// TIA Portal V20 export
TYPE "Stationsvariablen"
   STRUCT
      Anwahl_Tipp : Bool := FALSE;
      Status_Anw : Bool := FALSE;
      Anwahl_GS : Bool := FALSE;
      Status_GS : Bool;
      Status_Sicher : Bool;
      Tipp_Plus : Bool := FALSE;
      LEER : Bool := FALSE;
      Vorhanden : Bool := FALSE;
      IO : Bool := FALSE;
      NIO : Bool := FALSE;
      Reset_Teilestatus : Bool;
      Manu_Freigabe_SK : Bool;
      Richten_lauft : Bool;
      SNr : Int := 0;
      SK_Fertig : Bool;
      Taktzeit_max_Störung : Bool;
      Reserve_Einzelschritt : Array[0..31] of Bool;
   END_STRUCT;
   // Reserve_Einzelschritt[0..31] := FALSE;
END_TYPE
